FUNCTION_BLOCK Waypoint (* CAT Function Block Type *)
  (* Standard: 61499-2 *)
  (* Version 0.0, 7/9/2026, template *)
  PACKAGE Main;
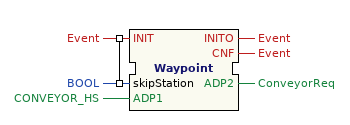
  EVENT_INPUT
    INIT WITH skipStation; (* Initialization Request *)
  END_EVENT
  EVENT_OUTPUT
    INITO; (* Initialization Confirm *)
    CNF; (* Execution Confirmation *)
  END_EVENT
  VAR_INPUT
    skipStation : BOOL; (* Input event qualifier *)
  END_VAR
  SOCKETS
    ADP1 : CONVEYOR_HS;
  END_SOCKETS
  PLUGS
    ADP2 : ConveyorReq;
  END_PLUGS
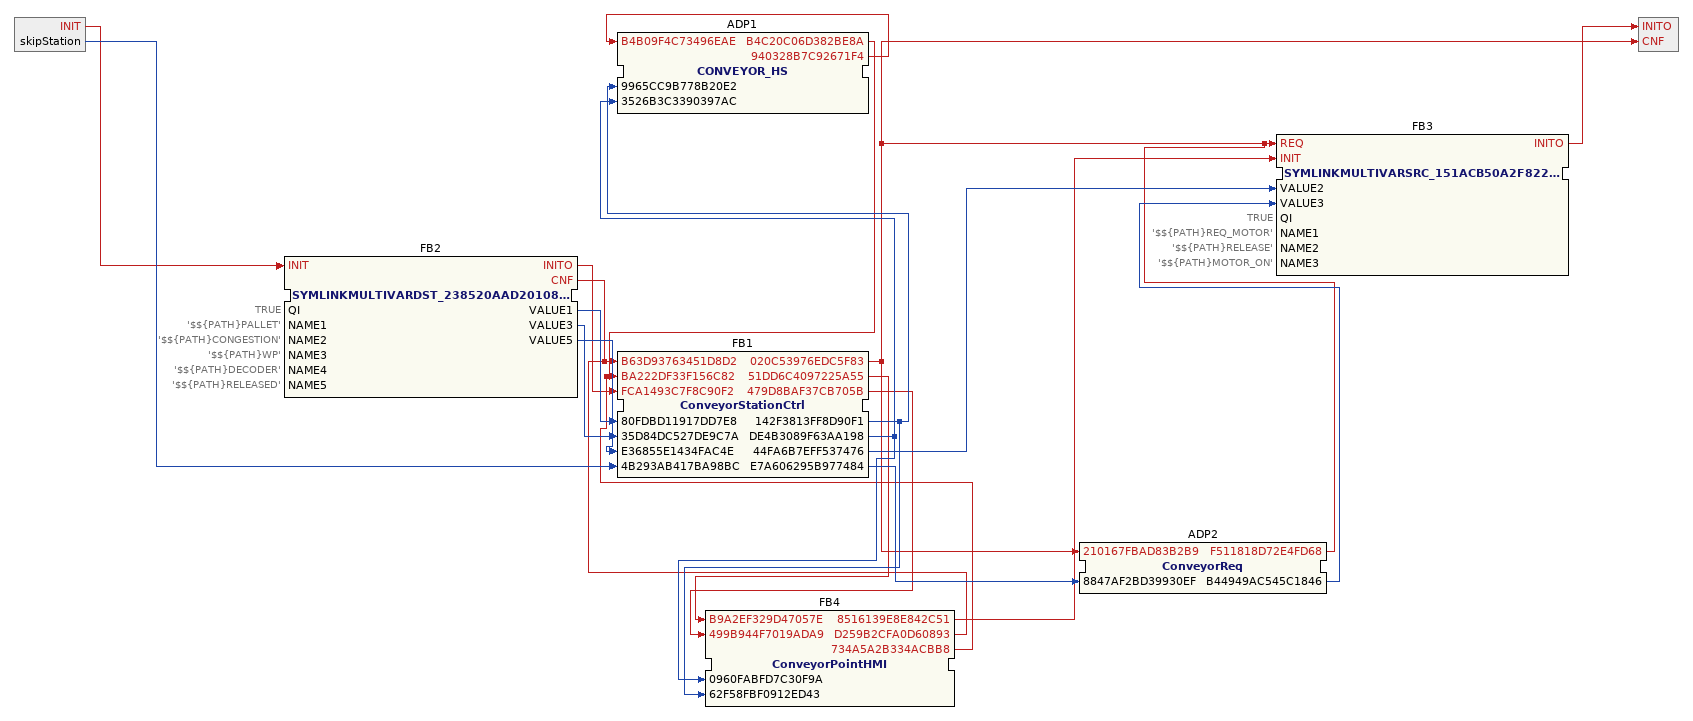
  FBS
    FB1 : ConveyorStationCtrl;
    FB2 : SYMLINKMULTIVARDST_238520AAD20108C65(QI := TRUE, NAME1 := '$${PATH}PALLET', NAME2 := '$${PATH}CONGESTION', NAME3 := '$${PATH}WP', NAME4 := '$${PATH}DECODER', NAME5 := '$${PATH}RELEASED'); {SET_ATTRIBUTE(Configuration.GenericFBType.InterfaceParams, Runtime.System#I:=7;VALUE${I$}:BOOL,BOOL,BOOL,BOOL,BOOL,BOOL,BOOL)}
    FB3 : SYMLINKMULTIVARSRC_151ACB50A2F8223B2(QI := TRUE, NAME1 := '$${PATH}REQ_MOTOR', NAME2 := '$${PATH}RELEASE', NAME3 := '$${PATH}MOTOR_ON'); {SET_ATTRIBUTE(Configuration.GenericFBType.InterfaceParams, Runtime.System#I:=3;VALUE${I$}:BOOL,BOOL,BOOL)}
    FB4 : ConveyorPointHMI;
  END_FBS
  EVENT_CONNECTIONS
    INIT TO FB2.INIT;
    FB3.INITO TO INITO;
    FB1.020C53976EDC5F83 TO CNF;
    FB1.020C53976EDC5F83 TO ADP2.210167FBAD83B2B9;
    FB1.020C53976EDC5F83 TO FB3.REQ;
    ADP2.F511818D72E4FD68 TO FB3.REQ;
    FB4.8516139E8E842C51 TO FB3.INIT;
    FB1.51DD6C4097225A55 TO FB4.B9A2EF329D47057E;
    FB1.479D8BAF37CB705B TO FB4.499B944F7019ADA9;
    FB4.D259B2CFA0D60893 TO FB1.B63D93763451D8D2;
    FB4.734A5A2B334ACBB8 TO FB1.BA222DF33F156C82;
    FB2.INITO TO FB1.FCA1493C7F8C90F2;
    FB2.CNF TO FB1.B63D93763451D8D2;
    ADP1.B4C20C06D382BE8A TO FB1.BA222DF33F156C82;
    ADP1.940328B7C92671F4 TO ADP1.B4B09F4C73496EAE;
  END_CONNECTIONS
  DATA_CONNECTIONS
    FB2.VALUE1 TO FB1.80FDBD11917DD7E8;
    FB2.VALUE3 TO FB1.35D84DC527DE9C7A;
    FB2.VALUE5 TO FB1.E36855E1434FAC4E;
    skipStation TO FB1.4B293AB417BA98BC;
    FB1.142F3813FF8D90F1 TO ADP1.9965CC9B778B20E2;
    FB1.DE4B3089F63AA198 TO ADP1.3526B3C3390397AC;
    FB1.44FA6B7EFF537476 TO FB3.VALUE2;
    FB1.E7A606295B977484 TO ADP2.8847AF2BD39930EF;
    FB1.DE4B3089F63AA198 TO FB4.0960FABFD7C30F9A;
    FB1.142F3813FF8D90F1 TO FB4.62F58FBF0912ED43;
    ADP2.B44949AC545C1846 TO FB3.VALUE3;
  END_CONNECTIONS
END_FUNCTION_BLOCK
